(* IEC 61131-3 sources: JingjiangArm/moonboxpro_arm_8.4/Application/Application/数据类型/系统参数/其他参数集, 9 files *)

(* ---- StArc_Mol_Param.st ---- *)
(*@CES
Name=StArc_Mol_Param
Type=Gvl
TypeGuid=2db5746d-d284-4425-9f7f-2663a34b0ebc
Guid=fa3e3698-9f51-498f-bb40-b12e90f03388
HasDeclaration=True
HasImplementation=False
*)
{DECLARATION}
{attribute 'pack_mode' := '1'}
(*2025.3.5.143340||35BYTES*)
TYPE StArc_Mol_Param :
STRUCT
	xUse_NewArcMol							: BOOL;(*给新算法先加个开关，后续可能不用了-先2025.3.5.152830*)
	(*2025.3.5.143328+*)
	(*套色模型计算pid函数获取的pid值@Cal_Kp_Ki|30bytes*)
	xUsePID_Mol								: BOOL;(*使用标志@代码中未用该变量,先留着吧*)
	rKadj_PID_Mol							: REAL;(*模型的pid增益_初始增益@开机和接料使用*)
	rKadj_I_Mol								: REAL;(*模型的I值增益_初始增益@开机和接料使用*)
	rKp_MolCal								: REAL;
	rKi_MolCal								: REAL;
	(*2024.9.2.083021 增加稳态和接料的模型参数*)
	byKadj_SetType							: BYTE;(*套色K值设置方式@ =0|使用初始增益|=1根据状态设置*)(*2024.9.2.131145 使用扩展参数种*)
	byArcAdjSts								: BYTE;(*套色调整状态@=0 初始状态(增益略大) |=1 稳态状态(增益略小)*)
	rKadj_PID_Mol_SteadySts					: REAL;(*模型的pid增益_稳态增益*)
	rKadj_I_Mol_SteadySts					: REAL;(*模型的I值增益_稳态增益*)
	(*2025.1.11.174053@v3方式的幅值裕度和相位裕度*)
	rMargin_Mag_Arc							: REAL:=20;
	rMargin_Phi_Arc							: REAL:=50;

(*套色陷波器*)
	xUseAntiNotch_Arc			: BOOL;(*套色使用陷波器@*)
	rWn_Arc						: REAL;(*陷波中心频率 rad/s*)
	rBw_Arc						: REAL;(*陷波宽度 rad/s*)
	rDp_Arc						: REAL;(*陷波深度 dB*)

	xUsePeriodic				: BOOL;(*使用Periodic方法*)
	rG_Periodic					: REAL;(*趋近增益  不同频率可能符号改变*)
	rW_Periodic					: REAL;(*需要抑制的频率，应该尽可能精确*)

	stStArcSpeedUpParam										: StArcSpeedUp;(*套色升速模型参数@30bytes|双积分*)
	stStArcSpeedUpFeedforward								: StArcSpeedUpFeedforward;(*前馈参数@30bytes*)

	rKp_GC						: REAL;
	rKi_GC						: REAL;
	rKd_GC						: REAL;
	rN_GC						: REAL;
	xCompensateEn_H				: BOOL;
	byCompensateValue_Hor		: BYTE;
	byMaxAddValue_Total_Hor		: BYTE;
	(*2026.5.14.191903+ 小郭测试算法@8bytes*)
    rPM_deg    : REAL :=50;    (* 目标相位裕度 60->50q(*2026.05.21.220750||wang.xy*)(°) *)

    rWc_Ts     : REAL :=0.3;    (* 归一化穿越频率 *)

	abyReserved:ARRAY [1..4] OF BYTE;(*预留31个字节*)
					(*12-->4*)

END_STRUCT
END_TYPE

{IMPLEMENTATION}

(* ---- StArcSpeedUp.st ---- *)
(*@CES
Name=StArcSpeedUp
Type=Gvl
TypeGuid=2db5746d-d284-4425-9f7f-2663a34b0ebc
Guid=efa365e6-af1e-4d1e-a80c-1fadbf9c4286
HasDeclaration=True
HasImplementation=False
*)
{DECLARATION}
{attribute 'pack_mode' := '1'}
TYPE StArcSpeedUp :
(*套色升速参数@主要是小黄设计的双积分控制器的参数*)
(*每个轴的参数都可能不一样@30bytes*)
STRUCT
	rK:REAL;(*增益系数*)
	rA2:REAL;(*模型参数*)
	rA1:REAL;(*模型参数*)
	rA0:REAL;(*模型参数*)
	abyReserved:ARRAY [1..14] OF BYTE;
END_STRUCT
END_TYPE

{IMPLEMENTATION}

(* ---- StArcSpeedUpFeedforward.st ---- *)
(*@CES
Name=StArcSpeedUpFeedforward
Type=Gvl
TypeGuid=2db5746d-d284-4425-9f7f-2663a34b0ebc
Guid=b9193669-47b2-40da-89b1-6ca603c59eae
HasDeclaration=True
HasImplementation=False
*)
{DECLARATION}
{attribute 'pack_mode' := '1'}
TYPE StArcSpeedUpFeedforward :
(*套色升速前馈@30BYTES*)
STRUCT
	rK:REAL;(*前馈系数-低速段*)
	rK_2:REAL;(*前馈系数-高速段*)
	abyReserved:ARRAY [1..22] OF BYTE;
(*	abyReserved:ARRAY [1..26] OF BYTE;*)
END_STRUCT
END_TYPE
{IMPLEMENTATION}

(* ---- StAxisCfgStruct.st ---- *)
(*@CES
Name=StAxisCfgStruct
Type=Gvl
TypeGuid=2db5746d-d284-4425-9f7f-2663a34b0ebc
Guid=69d05dad-9768-48d4-85b0-14945c9a532b
HasDeclaration=True
HasImplementation=False
*)
{DECLARATION}
{attribute 'pack_mode' := '1'}
TYPE StAxisCfgStruct :
STRUCT
	dwAxisProf		: DWORD:= 0;
							(*
							/ bit0=TRUE 轴打开
							/ bit1=TRUE 运动反向
							/ bit2=TRUE 采样反向()
							/ bit3~bit30 保留
							/ bit31=TRUE 站点存在于列表中
							*)
	iSid			: INT:= -1;
							(*
							/ -1表示无效轴
							/ 1~255(采用GNS方案后0作为GNS的默认分配/不体现在系统配置中
							*)
	iUnitId          :INT:=1;
END_STRUCT
END_TYPE

{IMPLEMENTATION}

(* ---- StMechanicalParamBuf.st ---- *)
(*@CES
Name=StMechanicalParamBuf
Type=Gvl
TypeGuid=2db5746d-d284-4425-9f7f-2663a34b0ebc
Guid=fd3f6fab-ce8b-4859-9675-c32c92772a95
HasDeclaration=True
HasImplementation=False
*)
{DECLARATION}
{attribute 'pack_mode' := '1'}
TYPE StMechanicalParamBuf :
STRUCT
	abyBuf	: ARRAY [1..200] OF BYTE;
END_STRUCT
END_TYPE

{IMPLEMENTATION}

(* ---- StStdVolParam_DnCut_UpCut.st ---- *)
(*@CES
Name=StStdVolParam_DnCut_UpCut
Type=Gvl
TypeGuid=2db5746d-d284-4425-9f7f-2663a34b0ebc
Guid=0efb4f92-3457-447a-bc79-dd669d3876a7
HasDeclaration=True
HasImplementation=False
*)
{DECLARATION}
{attribute 'pack_mode' := '1'}
TYPE StStdVolParam_DnCut_UpCut :
STRUCT
	alrStdVol_Diam		: ARRAY [1..4] OF LREAL;(* 标准卷径值 *)
	alrStdVol_Volt_AxisA: ARRAY [1..4] OF LREAL; (* 标准卷径对应的电压值|2019.1.25.142552|更名A轴 *)
	alrStdVol_Coef_AxisA: ARRAY [0..4] OF LREAL; (* 分段系数|2019.1.25.142601|更名A轴|[0]表<=1,[1]表>1&& <=2,[2]表>2&& <=3,[3]表>3&& <=4,[4]表>4 *)
	alrStdVol_Volt_AxisB: ARRAY [1..4] OF LREAL; (* 标准卷径对应的电压值|2019.1.25.142524|新增B轴 *)
	alrStdVol_Coef_AxisB: ARRAY [0..4] OF LREAL; (* 分段系数|2019.1.25.142542|新增B轴|[0]表<=1,[1]表>1&& <=2,[2]表>2&& <=3,[3]表>3&& <=4,[4]表>4 *)
	abyReserved: ARRAY [1..50] OF BYTE; (* 保留区域 *)
END_STRUCT
END_TYPE

{IMPLEMENTATION}

(* ---- StSysCfgStruct.st ---- *)
(*@CES
Name=StSysCfgStruct
Type=Gvl
TypeGuid=2db5746d-d284-4425-9f7f-2663a34b0ebc
Guid=08cdf89d-7f9f-4b4a-ba7e-4b606e266345
HasDeclaration=True
HasImplementation=False
*)
{DECLARATION}
{attribute 'pack_mode' := '1'}
TYPE StSysCfgStruct :
STRUCT
	iCompanyId					: INT := 0;(* 公司id/0科赛/1飞达/... *)
	byLanguageId				: BYTE := 1;(* 语言id/1.中文/2.英文/... *)
	byUnitMaxNum				: BYTE := 7;(* 色组数量/0~MAX_UNIT_NUM *)
	astStAxisCfgStruct_UW_I		: ARRAY [1..2] OF StAxisCfgStruct;(* UW: UnWind/放料 *)
	astStAxisCfgStruct_RW_I		: ARRAY [1..2] OF StAxisCfgStruct;(* RW: ReWind/收料 *)
	stStAxisCfgStruct_IF_I		: StAxisCfgStruct;(* IF: InFeed/放牵 *)
	stStAxisCfgStruct_OF_I		: StAxisCfgStruct;(* OF: OutFeed/收牵 *)
	astStAxisCfgStruct_CD_I		: ARRAY [1..2] OF StAxisCfgStruct;(* CD: Central Drum/中心滚筒 *)(*中心辊增加一个|2024.04.01.094732*)
	astStAxisCfgStruct_UW_II		: ARRAY [1..2] OF StAxisCfgStruct;(* UW: UnWind/放料 *)
	astStAxisCfgStruct_RW_II		: ARRAY [1..2] OF StAxisCfgStruct;(* RW: ReWind/收料 *)
	stStAxisCfgStruct_IF_II		: StAxisCfgStruct;(* IF: InFeed/放牵 *)
	stStAxisCfgStruct_OF_II		: StAxisCfgStruct;(* OF: OutFeed/收牵 *)
	astStAxisCfgStruct_CD_II		: ARRAY [1..2] OF StAxisCfgStruct;(* CD: Central Drum/中心滚筒 *)(*中心辊增加一个|2024.04.01.094732*)

	astStAxisCfgStruct_PC_		: ARRAY [1..MAX_UNIT_NUM] OF StAxisCfgStruct;(*光电眼行走机构 | 2024.04.01.092649*)
	astStAxisCfgStruct_BR_		: ARRAY [1..MAX_UNIT_NUM] OF StAxisCfgStruct;(* BR: Bottom Roller/底辊 *)
	astStAxisCfgStruct_PR_		: ARRAY [1..MAX_UNIT_NUM] OF StAxisCfgStruct;(* PR: Prn Roller/版辊 *)
	astStAxisCfgStruct_NR_		: ARRAY [1..MAX_UNIT_NUM] OF StAxisCfgStruct;(* NR: Net Roller/网辊 *)
	astStAxisCfgStruct_PR_M_	: ARRAY [1..MAX_UNIT_NUM] OF StAxisCfgStruct;(* PR_M: PrnRoller Mside/版辊压力M侧 *)
	astStAxisCfgStruct_PR_G_	: ARRAY [1..MAX_UNIT_NUM] OF StAxisCfgStruct;(* PR_G: PrnRoller Gside/版辊压力G侧 *)
	astStAxisCfgStruct_NR_M_	: ARRAY [1..MAX_UNIT_NUM] OF StAxisCfgStruct;(* NR_M: NetRoller Mside/网辊压力M侧 *)
	astStAxisCfgStruct_NR_G_	: ARRAY [1..MAX_UNIT_NUM] OF StAxisCfgStruct;(* NR_G: NetRoller Gside/网辊压力G侧 *)
	astStAxisCfgStruct_STR_M_	: ARRAY [1..MAX_UNIT_NUM] OF StAxisCfgStruct;(* NR_M: NetRoller Mside/张带辊压力M侧 *)
	astStAxisCfgStruct_STR_G_	: ARRAY [1..MAX_UNIT_NUM] OF StAxisCfgStruct;(* NR_G: NetRoller Gside/张带辊压力G侧 *)
	astStAxisCfgStruct_HORIZ_	: ARRAY [1..MAX_UNIT_NUM] OF StAxisCfgStruct;(* HORIZ: 横向控制电机 *)
//系统配置参数内容更新，记得重新保存
	astStAxisCfgStruct_Ctl_	: ARRAY [1..MAX_UNIT_NUM] OF StAxisCfgStruct;(* HORIZ: 横向控制电机 *)

END_STRUCT
END_TYPE

{IMPLEMENTATION}

(* ---- StTimeSet_DnCut_UpCut.st ---- *)
(*@CES
Name=StTimeSet_DnCut_UpCut
Type=Gvl
TypeGuid=2db5746d-d284-4425-9f7f-2663a34b0ebc
Guid=3d90f000-d022-493a-8845-04f294dfa37c
HasDeclaration=True
HasImplementation=False
*)
{DECLARATION}
{attribute 'pack_mode' := '1'}
TYPE StTimeSet_DnCut_UpCut :
STRUCT
	iDelayMsec_CutterHolder			: INT; (* 裁刀架延时 *)
	iDelayMsec_RollerCylinder		: INT; (* 胶辊汽缸延时 *)
	iDelayMsec_CutOffKnifeCylinder	: INT; (* 裁刀汽缸延时 *)
	uiMM_Roller2GummedTape			: UINT; (* 压辊压在料上距胶带的距离/单位:mm *)
	uiMM_Roller2CutOfKnife			: UINT; (* 压辊距裁刀的材料距离|单位:mm *)
	uiMM_CutOfKnife2GummedTape		: UINT; (* 裁刀距胶带的距离/单位:mm *)
	iStepVariation4ChangeTime		: INT; (* 2018.9.30.100457/用来步进胶辊延时和裁刀延时的变化量 *)
	iDelaySec_AirInflation_Mixed	: INT; (* 一刀双裁大臂充气延时/2019.6.20.175319 *)
	iHodTime_HelpStep_RollerCylinder: INT;(*2021.7.17.140936 增加接料压辊助走持续时间--ALTMA*)
	rStepVariation4ChangeDis		: REAL;(*参考距离值|2022.10.13.105318|mm*)
	abyRsvdFields						: ARRAY [1..44] OF BYTE; (* 保留区域 *)
	(*2022.10.13.105336 +rStepVariation4ChangeDis|48-->44*)
END_STRUCT
END_TYPE

{IMPLEMENTATION}

(* ---- StVarList.st ---- *)
(*@CES
Name=StVarList
Type=Gvl
TypeGuid=2db5746d-d284-4425-9f7f-2663a34b0ebc
Guid=8fe36071-a98d-4a3e-9449-8cd49bd30799
HasDeclaration=True
HasImplementation=False
*)
{DECLARATION}
{attribute 'pack_mode' := '1'}
//xi.hy新增@七号以后
TYPE StVarList:
STRUCT
	wVirTual_Cnt:WORD;//虚拟码盘计数
	wVirTual_Sts:WORD;//虚拟码盘状态
	dwTime_Lock:DWORD;//锁存时间
	dwEnc_Lock:DWORD;//锁存编码器
END_STRUCT
END_TYPE

{IMPLEMENTATION}
